(* IEC 61131-3 sources: codesys-framework/txt/application/ToDo/Hardware/IO/Camera, 3 files *)

(* ---- E_CameraStates.dut.st ---- *)
{attribute 'qualified_only'}
{attribute 'strict'}
TYPE E_CameraStates :
(
	Invalid := 0,
	None,
	Initialize,
	Connect,
	Disconnect,
	Standby,
	SelectJob,
	TakePicture,
	Reset
);
END_TYPE

(* ---- SC_SystemParametersVisuCamera.dut.st ---- *)
TYPE SC_SystemParametersVisuCamera :
STRUCT
	adress 			: NBS.IP_ADDR;
	conTimeout 		: UDINT;
	readPort 		: UINT;
	writePort 		: UINT;
	cycleTime 		: TIME;
	monitorTime 	: TIME;
	shutterTime 	: TIME;
	readTimeout 	: TIME;
	jobTimeout 		: TIME;
END_STRUCT
END_TYPE

(* ---- FB_Camera.pou.st ---- *)
FUNCTION_BLOCK FB_Camera IMPLEMENTS I_Camera
VAR_INPUT
END_VAR
VAR_OUTPUT
END_VAR
VAR
	_scSysPar 				: SC_SystemParametersVisuCamera;

	_eState 				: E_CameraStates;
	_xBusy 					: BOOL;
	_xDone 					: BOOL;
	_xError 				: BOOL;
	_iErrorId 				: UINT;
	_sError 				: STRING;

	_read 	  				: NBS.TCP_Read;
	_write		 			: NBS.TCP_Write;
	_writeFeedBack 			: NBS.TCP_Read;

	_clientState			: NBS.TCP_Client;
	_clientRead        		: NBS.TCP_Client;
	_clientWrite			: NBS.TCP_Client;

	_tonMonitor 			: TON;
	_tonPicture 			: TON;
	_tonSelectJob 			: TON;

	_xConnected 			: BOOL;

	_iStateMonitor 			: UINT;
	_iStateConnect 			: UINT;
	_iStateSetJob 			: UINT;
	_iStateTakePicture 		: UINT;
	_iStateConnectMethod 	: UINT;
	_iStateDisconnect 		: UINT;

	_sJob 					: STRING;
	_sPicture 				: STRING;
	_sFeedBack 				: STRING;
	_id 					: UINT;

	_sResult 				: STRING(280);
	_sResultPrev			: STRING(280);
	_sPictureId				: STRING;
END_VAR

// --- BEGIN IMPLEMENTATION ---

Monitor();

ProcessFBs();
ProcessState();
